(* Schneider Machine Expert - Basic project modbus_03_read_q_fc1, file version 3.0.0.0 *)
(* ProjectInformations: Name=New project *)

HARDWARE
  Cpu 0: TM200CE40T
  EthernetConfiguration: NetworkName=M200, IpAllocationMode=FixedAddress, IpAddress=0.0.0.0, SubnetMask=0.0.0.0
  SerialLineConfiguration: Baud=Baud19200, Parity=ParityEven, DataBits=DataBits8, StopBits=StopBits1, PhysicalMedium=PhysicalMediumRs485, TransmissionMode=TransmissionModeModbusRtu, SlaveId=1, Addressing=MasterAddressing
  MastTask: UsePeriodScanMode=false, PeriodScan=100
  FastTask: Period=255
  CpuBehavior: StartingMode=StartAsPreviousState, AutoSaveRamOnEeprom=true, WatchdogPeriod=250

SYMBOLS  (address, symbol, comment, settings)
  %READ_VAR0   [Link(Value(FBComLinkParameterEnums=SerialLine1)), RemoteDeviceId(Value(int=1)), Timeout(Value(int=100)), ObjType(Value(FBComObjTypeParameterEnums=Q)), FirstObj(Value(int=41)), Quantity(Value(int=17)), IndexData(Value(int=220))]

POU Generated C++ - EXPERIMENTAL
  (* SectionNumber=0 *)

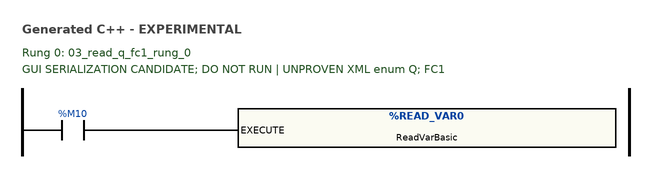

// Rung 0: 03_read_q_fc1_rung_0
// GUI SERIALIZATION CANDIDATE; DO NOT RUN | UNPROVEN XML enum Q; FC1
  BLK %READ_VAR0
  LD %M10
  EXECUTE
  END_BLK
  // as ST:
  //   %READ_VAR0(EXECUTE := %M10);
